{attribute 'qualified_only'}
VAR_GLOBAL CONSTANT
  DIRECTORY : T_MaxString := 'C:\TcUnit_IntecreFile';
  TIMEOUT : TIME := T#5S;
END_VAR

(* stored: Version 1.1.0.1, ProductVersion 3.1.4026.25
   GVL TestFiles: Id {aafe6cc2-d75f-402e-9e36-08d5a8212fc8} *)
